(* IEC 61131-3 sources: sceptre-phenix-topologies/cherrymountain-brewery/plant/generated/fleet/fr/openplc/fr-plc-cellar, 1 file *)

(* ---- located_vars.st ---- *)
(* Generated by plantgen from plant/plant.yaml and plant/sites.yaml (site fr). Do not edit. *)
(* Analog values are raw registers: engineering value = raw / 10^scaling. *)
(* RIO I/O is at %IX100.0 / %QX100.0 / %IW100 / %QW100 (v3 and v4 alike). *)
(* PLC memory: bits from %QX0.0 (coils), words from %MW0 (holding register qw_count and up, see modbus_slave.json). *)
VAR
  CEL_CLK_KI01_PV AT %IW100 : UINT; (* Cellar simulation clock (compressed fermentation time), h, x10 *)
  CEL_FV101_TT01_PV AT %IW101 : UINT; (* FV-101 side temperature, degF, x100 *)
  CEL_FV101_TT01_ALM_DEVIATION AT %QX0.0 : BOOL; (* FV-101 side temperature: deviation alarm (high) *)
  CEL_FV101_TT01_ALM_HIGH AT %QX0.1 : BOOL; (* FV-101 side temperature: high alarm (medium) *)
  CEL_FV101_TV01_CMD AT %QX100.0 : BOOL; (* FV-101 side glycol valve command *)
  CEL_FV101_TT02_PV AT %IW102 : UINT; (* FV-101 cone temperature, degF, x100 *)
  CEL_FV101_TT02_ALM_DEVIATION AT %QX0.2 : BOOL; (* FV-101 cone temperature: deviation alarm (medium) *)
  CEL_FV101_TV02_CMD AT %QX100.1 : BOOL; (* FV-101 cone glycol valve command *)
  CEL_FV101_PT01_PV AT %IW103 : UINT; (* FV-101 head pressure (absolute), psia, x100 *)
  CEL_FV101_PT01_ALM_HIGH AT %QX0.3 : BOOL; (* FV-101 head pressure (absolute): high alarm (high) *)
  CEL_FV101_PT01_ALM_LOW AT %QX0.4 : BOOL; (* FV-101 head pressure (absolute): low alarm (low) *)
  CEL_FV101_DT01_PV AT %IW104 : UINT; (* FV-101 apparent extract (sample-port density meter), degP, x100 *)
  CEL_FV101_PCV01_SP AT %QW100 : UINT; (* FV-101 spunding valve setpoint (absolute), psia, x100 *)
  CEL_FV101_ZSO01_PV AT %IX100.0 : BOOL; (* FV-101 spunding valve open (venting) *)
  CEL_FV101_TT01_SP AT %MW0 : UINT; (* FV-101 side temperature setpoint, degF, x100 *)
  CEL_FV101_TT02_SP AT %MW1 : UINT; (* FV-101 cone temperature setpoint, degF, x100 *)
  CEL_FV102_TT01_PV AT %IW105 : UINT; (* FV-102 side temperature, degF, x100 *)
  CEL_FV102_TT01_ALM_DEVIATION AT %QX0.5 : BOOL; (* FV-102 side temperature: deviation alarm (high) *)
  CEL_FV102_TT01_ALM_HIGH AT %QX0.6 : BOOL; (* FV-102 side temperature: high alarm (medium) *)
  CEL_FV102_TV01_CMD AT %QX100.2 : BOOL; (* FV-102 side glycol valve command *)
  CEL_FV102_TT02_PV AT %IW106 : UINT; (* FV-102 cone temperature, degF, x100 *)
  CEL_FV102_TT02_ALM_DEVIATION AT %QX0.7 : BOOL; (* FV-102 cone temperature: deviation alarm (medium) *)
  CEL_FV102_TV02_CMD AT %QX100.3 : BOOL; (* FV-102 cone glycol valve command *)
  CEL_FV102_PT01_PV AT %IW107 : UINT; (* FV-102 head pressure (absolute), psia, x100 *)
  CEL_FV102_PT01_ALM_HIGH AT %QX1.0 : BOOL; (* FV-102 head pressure (absolute): high alarm (high) *)
  CEL_FV102_PT01_ALM_LOW AT %QX1.1 : BOOL; (* FV-102 head pressure (absolute): low alarm (low) *)
  CEL_FV102_DT01_PV AT %IW108 : UINT; (* FV-102 apparent extract (sample-port density meter), degP, x100 *)
  CEL_FV102_PCV01_SP AT %QW101 : UINT; (* FV-102 spunding valve setpoint (absolute), psia, x100 *)
  CEL_FV102_ZSO01_PV AT %IX100.1 : BOOL; (* FV-102 spunding valve open (venting) *)
  CEL_FV102_TT01_SP AT %MW2 : UINT; (* FV-102 side temperature setpoint, degF, x100 *)
  CEL_FV102_TT02_SP AT %MW3 : UINT; (* FV-102 cone temperature setpoint, degF, x100 *)
  CEL_FV103_TT01_PV AT %IW109 : UINT; (* FV-103 side temperature, degF, x100 *)
  CEL_FV103_TT01_ALM_DEVIATION AT %QX1.2 : BOOL; (* FV-103 side temperature: deviation alarm (high) *)
  CEL_FV103_TT01_ALM_HIGH AT %QX1.3 : BOOL; (* FV-103 side temperature: high alarm (medium) *)
  CEL_FV103_TV01_CMD AT %QX100.4 : BOOL; (* FV-103 side glycol valve command *)
  CEL_FV103_TT02_PV AT %IW110 : UINT; (* FV-103 cone temperature, degF, x100 *)
  CEL_FV103_TT02_ALM_DEVIATION AT %QX1.4 : BOOL; (* FV-103 cone temperature: deviation alarm (medium) *)
  CEL_FV103_TV02_CMD AT %QX100.5 : BOOL; (* FV-103 cone glycol valve command *)
  CEL_FV103_PT01_PV AT %IW111 : UINT; (* FV-103 head pressure (absolute), psia, x100 *)
  CEL_FV103_PT01_ALM_HIGH AT %QX1.5 : BOOL; (* FV-103 head pressure (absolute): high alarm (high) *)
  CEL_FV103_PT01_ALM_LOW AT %QX1.6 : BOOL; (* FV-103 head pressure (absolute): low alarm (low) *)
  CEL_FV103_DT01_PV AT %IW112 : UINT; (* FV-103 apparent extract (sample-port density meter), degP, x100 *)
  CEL_FV103_PCV01_SP AT %QW102 : UINT; (* FV-103 spunding valve setpoint (absolute), psia, x100 *)
  CEL_FV103_ZSO01_PV AT %IX100.2 : BOOL; (* FV-103 spunding valve open (venting) *)
  CEL_FV103_TT01_SP AT %MW4 : UINT; (* FV-103 side temperature setpoint, degF, x100 *)
  CEL_FV103_TT02_SP AT %MW5 : UINT; (* FV-103 cone temperature setpoint, degF, x100 *)
  CEL_FV104_TT01_PV AT %IW113 : UINT; (* FV-104 side temperature, degF, x100 *)
  CEL_FV104_TT01_ALM_DEVIATION AT %QX1.7 : BOOL; (* FV-104 side temperature: deviation alarm (high) *)
  CEL_FV104_TT01_ALM_HIGH AT %QX2.0 : BOOL; (* FV-104 side temperature: high alarm (medium) *)
  CEL_FV104_TV01_CMD AT %QX100.6 : BOOL; (* FV-104 side glycol valve command *)
  CEL_FV104_TT02_PV AT %IW114 : UINT; (* FV-104 cone temperature, degF, x100 *)
  CEL_FV104_TT02_ALM_DEVIATION AT %QX2.1 : BOOL; (* FV-104 cone temperature: deviation alarm (medium) *)
  CEL_FV104_TV02_CMD AT %QX100.7 : BOOL; (* FV-104 cone glycol valve command *)
  CEL_FV104_PT01_PV AT %IW115 : UINT; (* FV-104 head pressure (absolute), psia, x100 *)
  CEL_FV104_PT01_ALM_HIGH AT %QX2.2 : BOOL; (* FV-104 head pressure (absolute): high alarm (high) *)
  CEL_FV104_PT01_ALM_LOW AT %QX2.3 : BOOL; (* FV-104 head pressure (absolute): low alarm (low) *)
  CEL_FV104_DT01_PV AT %IW116 : UINT; (* FV-104 apparent extract (sample-port density meter), degP, x100 *)
  CEL_FV104_PCV01_SP AT %QW103 : UINT; (* FV-104 spunding valve setpoint (absolute), psia, x100 *)
  CEL_FV104_ZSO01_PV AT %IX100.3 : BOOL; (* FV-104 spunding valve open (venting) *)
  CEL_FV104_TT01_SP AT %MW6 : UINT; (* FV-104 side temperature setpoint, degF, x100 *)
  CEL_FV104_TT02_SP AT %MW7 : UINT; (* FV-104 cone temperature setpoint, degF, x100 *)
  CEL_BBT201_TT01_PV AT %IW117 : UINT; (* BBT-201 temperature, degF, x100 *)
  CEL_BBT201_TT01_ALM_DEVIATION AT %QX2.4 : BOOL; (* BBT-201 temperature: deviation alarm (medium) *)
  CEL_BBT201_PT01_PV AT %IW118 : UINT; (* BBT-201 head pressure (absolute), psia, x100 *)
  CEL_BBT201_PT01_ALM_HIGH AT %QX2.5 : BOOL; (* BBT-201 head pressure (absolute): high alarm (high) *)
  CEL_BBT201_LT01_PV AT %IW119 : UINT; (* BBT-201 level, %, x10 *)
  CEL_BBT201_AT01_PV AT %IW120 : UINT; (* BBT-201 dissolved CO2 (inline meter), vol, x100 *)
  CEL_BBT201_FT01_PV AT %IW121 : UINT; (* BBT-201 carbonation stone CO2 flow, L/min, x10 *)
  CEL_BBT201_TV01_CMD AT %QX101.0 : BOOL; (* BBT-201 jacket glycol valve command *)
  CEL_BBT201_XV01_CMD AT %QX101.1 : BOOL; (* BBT-201 outlet valve (to packaging) *)
  CEL_BBT201_FCV01_OUT AT %QW104 : UINT; (* BBT-201 carbonation CO2 flow valve position, %, x10 *)
  CEL_BBT201_TT01_SP AT %MW8 : UINT; (* BBT-201 temperature setpoint, degF, x100 *)
  CEL_BBT201_AT01_SP AT %MW9 : UINT; (* BBT-201 carbonation target, vol, x100 *)
  CEL_BBT201_PT01_SP AT %MW10 : UINT; (* BBT-201 equilibrium head pressure for the target (computed, absolute), psia, x100 *)
  CEL_BBT202_TT01_PV AT %IW122 : UINT; (* BBT-202 temperature, degF, x100 *)
  CEL_BBT202_TT01_ALM_DEVIATION AT %QX2.6 : BOOL; (* BBT-202 temperature: deviation alarm (medium) *)
  CEL_BBT202_PT01_PV AT %IW123 : UINT; (* BBT-202 head pressure (absolute), psia, x100 *)
  CEL_BBT202_PT01_ALM_HIGH AT %QX2.7 : BOOL; (* BBT-202 head pressure (absolute): high alarm (high) *)
  CEL_BBT202_LT01_PV AT %IW124 : UINT; (* BBT-202 level, %, x10 *)
  CEL_BBT202_AT01_PV AT %IW125 : UINT; (* BBT-202 dissolved CO2 (inline meter), vol, x100 *)
  CEL_BBT202_FT01_PV AT %IW126 : UINT; (* BBT-202 carbonation stone CO2 flow, L/min, x10 *)
  CEL_BBT202_TV01_CMD AT %QX101.2 : BOOL; (* BBT-202 jacket glycol valve command *)
  CEL_BBT202_XV01_CMD AT %QX101.3 : BOOL; (* BBT-202 outlet valve (to packaging) *)
  CEL_BBT202_FCV01_OUT AT %QW105 : UINT; (* BBT-202 carbonation CO2 flow valve position, %, x10 *)
  CEL_BBT202_TT01_SP AT %MW11 : UINT; (* BBT-202 temperature setpoint, degF, x100 *)
  CEL_BBT202_AT01_SP AT %MW12 : UINT; (* BBT-202 carbonation target, vol, x100 *)
  CEL_BBT202_PT01_SP AT %MW13 : UINT; (* BBT-202 equilibrium head pressure for the target (computed, absolute), psia, x100 *)
  CEL_DH_ZSC01_PV AT %IX100.4 : BOOL; (* Hop port closed *)
  CEL_DH_XV01_CMD AT %QX101.4 : BOOL; (* Hop port CO2 purge valve *)
  CEL_DH_XV02_CMD AT %QX101.5 : BOOL; (* Hop dose valve *)
  CEL_DH_XC01_CMD AT %QX3.0 : BOOL; (* Dry-hop dose request (operator; fr-plc-cellar purges, doses, and clears it) *)
  CEL_DH_XS01_STEP AT %MW14 : UINT; (* Dry-hop sequence step (0 idle, 1 CO2 purge, 2 dose), None, x1 *)
  CEL_XFER_ZS01_PV AT %IX100.5 : BOOL; (* Transfer route verified (swing-panel proximity) *)
  CEL_XFER_YS01_PV AT %IX100.6 : BOOL; (* Transfer pump running *)
  CEL_XFER_FT01_PV AT %IW127 : UINT; (* Transfer flow, gal/min, x10 *)
  CEL_XFER_HS01_CMD AT %QX101.6 : BOOL; (* Transfer pump run command *)
  CEL_XFER_XS01_ACTIVE AT %QX3.1 : BOOL; (* Transfer in progress (peer status for fr-plc-utilities) *)
  CEL_XFER_XS02_CIP_PERMIT AT %QX3.2 : BOOL; (* CIP permitted on the cellar circuits (peer status for fr-plc-utilities) *)
  CEL_SYS_XS01_CO2_OK AT %IX100.7 : BOOL; (* Cellar CO2 relay healthy (below 15,000 ppm, detection powered) *)
  CEL_SYS_XS01_CO2_INHIBIT AT %QX3.3 : BOOL; (* Carbonation inhibited by the cellar CO2 relay (fr-plc-cellar interlock) *)
  CEL_SYS_XS01_ALM_STATE AT %QX3.4 : BOOL; (* Carbonation inhibited by the cellar CO2 relay (fr-plc-cellar interlock): state alarm (medium) *)
  CEL_PSV_ZSH01_PV AT %IX101.0 : BOOL; (* FV-101 relief valve (PSV) lifted *)
  CEL_PSV_ZSH01_ALM_STATE AT %QX3.5 : BOOL; (* FV-101 relief valve (PSV) lifted: state alarm (high) *)
  CEL_PSV_ZSH02_PV AT %IX101.1 : BOOL; (* FV-102 relief valve (PSV) lifted *)
  CEL_PSV_ZSH02_ALM_STATE AT %QX3.6 : BOOL; (* FV-102 relief valve (PSV) lifted: state alarm (high) *)
  CEL_PSV_ZSH03_PV AT %IX101.2 : BOOL; (* FV-103 relief valve (PSV) lifted *)
  CEL_PSV_ZSH03_ALM_STATE AT %QX3.7 : BOOL; (* FV-103 relief valve (PSV) lifted: state alarm (high) *)
  CEL_PSV_ZSH04_PV AT %IX101.3 : BOOL; (* FV-104 relief valve (PSV) lifted *)
  CEL_PSV_ZSH04_ALM_STATE AT %QX4.0 : BOOL; (* FV-104 relief valve (PSV) lifted: state alarm (high) *)
  CEL_PSV_ZSH05_PV AT %IX101.4 : BOOL; (* BBT-201 relief valve (PSV) lifted *)
  CEL_PSV_ZSH05_ALM_STATE AT %QX4.1 : BOOL; (* BBT-201 relief valve (PSV) lifted: state alarm (high) *)
  CEL_PSV_ZSH06_PV AT %IX101.5 : BOOL; (* BBT-202 relief valve (PSV) lifted *)
  CEL_PSV_ZSH06_ALM_STATE AT %QX4.2 : BOOL; (* BBT-202 relief valve (PSV) lifted: state alarm (high) *)
  CEL_ENTRY_HS01_ENTRY AT %QX4.3 : BOOL; (* FV-101 entry permit issued (entry supervisor; locks the vessel out) *)
  CEL_ENTRY_HS02_ENTRY AT %QX4.4 : BOOL; (* FV-102 entry permit issued (entry supervisor; locks the vessel out) *)
  CEL_ENTRY_HS03_ENTRY AT %QX4.5 : BOOL; (* FV-103 entry permit issued (entry supervisor; locks the vessel out) *)
  CEL_ENTRY_HS04_ENTRY AT %QX4.6 : BOOL; (* FV-104 entry permit issued (entry supervisor; locks the vessel out) *)
  CEL_ENTRY_HS05_ENTRY AT %QX4.7 : BOOL; (* BBT-201 entry permit issued (entry supervisor; locks the vessel out) *)
  CEL_ENTRY_HS06_ENTRY AT %QX5.0 : BOOL; (* BBT-202 entry permit issued (entry supervisor; locks the vessel out) *)
  CEL_ENTRY_XS01_LOCKED AT %QX5.1 : BOOL; (* FV-101 locked out for entry (glycol, CO2, outlet, and CIP) *)
  CEL_ENTRY_XS02_LOCKED AT %QX5.2 : BOOL; (* FV-102 locked out for entry (glycol, CO2, outlet, and CIP) *)
  CEL_ENTRY_XS03_LOCKED AT %QX5.3 : BOOL; (* FV-103 locked out for entry (glycol, CO2, outlet, and CIP) *)
  CEL_ENTRY_XS04_LOCKED AT %QX5.4 : BOOL; (* FV-104 locked out for entry (glycol, CO2, outlet, and CIP) *)
  CEL_ENTRY_XS05_LOCKED AT %QX5.5 : BOOL; (* BBT-201 locked out for entry (glycol, CO2, outlet, and CIP) *)
  CEL_ENTRY_XS06_LOCKED AT %QX5.6 : BOOL; (* BBT-202 locked out for entry (glycol, CO2, outlet, and CIP) *)
  CEL_ENTRY_XS11_CIP_OK AT %QX5.7 : BOOL; (* FV-101 CIP permitted, not in entry (peer status for fr-plc-utilities) *)
  CEL_ENTRY_XS12_CIP_OK AT %QX6.0 : BOOL; (* FV-102 CIP permitted, not in entry (peer status for fr-plc-utilities) *)
  CEL_ENTRY_XS13_CIP_OK AT %QX6.1 : BOOL; (* FV-103 CIP permitted, not in entry (peer status for fr-plc-utilities) *)
  CEL_ENTRY_XS14_CIP_OK AT %QX6.2 : BOOL; (* FV-104 CIP permitted, not in entry (peer status for fr-plc-utilities) *)
  CEL_ENTRY_XS15_CIP_OK AT %QX6.3 : BOOL; (* BBT-201 CIP permitted, not in entry (peer status for fr-plc-utilities) *)
  CEL_ENTRY_XS16_CIP_OK AT %QX6.4 : BOOL; (* BBT-202 CIP permitted, not in entry (peer status for fr-plc-utilities) *)
  CEL_ENTRY_XA01_PV AT %QX6.5 : BOOL; (* FV-101 write to a locked-out valve during entry *)
  CEL_ENTRY_XA01_ALM_STATE AT %QX6.6 : BOOL; (* FV-101 write to a locked-out valve during entry: state alarm (critical) *)
  CEL_ENTRY_XA02_PV AT %QX6.7 : BOOL; (* FV-102 write to a locked-out valve during entry *)
  CEL_ENTRY_XA02_ALM_STATE AT %QX7.0 : BOOL; (* FV-102 write to a locked-out valve during entry: state alarm (critical) *)
  CEL_ENTRY_XA03_PV AT %QX7.1 : BOOL; (* FV-103 write to a locked-out valve during entry *)
  CEL_ENTRY_XA03_ALM_STATE AT %QX7.2 : BOOL; (* FV-103 write to a locked-out valve during entry: state alarm (critical) *)
  CEL_ENTRY_XA04_PV AT %QX7.3 : BOOL; (* FV-104 write to a locked-out valve during entry *)
  CEL_ENTRY_XA04_ALM_STATE AT %QX7.4 : BOOL; (* FV-104 write to a locked-out valve during entry: state alarm (critical) *)
  CEL_ENTRY_XA05_PV AT %QX7.5 : BOOL; (* BBT-201 write to a locked-out valve during entry *)
  CEL_ENTRY_XA05_ALM_STATE AT %QX7.6 : BOOL; (* BBT-201 write to a locked-out valve during entry: state alarm (critical) *)
  CEL_ENTRY_XA06_PV AT %QX7.7 : BOOL; (* BBT-202 write to a locked-out valve during entry *)
  CEL_ENTRY_XA06_ALM_STATE AT %QX8.0 : BOOL; (* BBT-202 write to a locked-out valve during entry: state alarm (critical) *)
  CEL_PROFILE_HS01_AUTO AT %QX8.1 : BOOL; (* FV-101 fermentation profile on (fr-plc-cellar sets its temperature setpoints) *)
  CEL_PROFILE_HS02_AUTO AT %QX8.2 : BOOL; (* FV-102 fermentation profile on (fr-plc-cellar sets its temperature setpoints) *)
  CEL_PROFILE_HS03_AUTO AT %QX8.3 : BOOL; (* FV-103 fermentation profile on (fr-plc-cellar sets its temperature setpoints) *)
  CEL_PROFILE_HS04_AUTO AT %QX8.4 : BOOL; (* FV-104 fermentation profile on (fr-plc-cellar sets its temperature setpoints) *)
  CEL_PROFILE_KS01_STAGE AT %MW15 : UINT; (* FV-101 profile stage (0 empty, 1 fermenting, 2 diacetyl rest, 3 crash), None, x1 *)
  CEL_PROFILE_KS02_STAGE AT %MW16 : UINT; (* FV-102 profile stage (0 empty, 1 fermenting, 2 diacetyl rest, 3 crash), None, x1 *)
  CEL_PROFILE_KS03_STAGE AT %MW17 : UINT; (* FV-103 profile stage (0 empty, 1 fermenting, 2 diacetyl rest, 3 crash), None, x1 *)
  CEL_PROFILE_KS04_STAGE AT %MW18 : UINT; (* FV-104 profile stage (0 empty, 1 fermenting, 2 diacetyl rest, 3 crash), None, x1 *)
  CEL_PROFILE_TC01_SP AT %MW19 : UINT; (* Profile temperature while the beer ferments, degF, x100 *)
  CEL_PROFILE_TC02_SP AT %MW20 : UINT; (* Profile temperature of the diacetyl rest, degF, x100 *)
  CEL_PROFILE_TC03_SP AT %MW21 : UINT; (* Profile temperature of the crash, degF, x100 *)
  CEL_PROFILE_KC01_SP AT %MW22 : UINT; (* Diacetyl rest length in plant minutes (180 is 144 h of fermentation on the range's 48x clock), min, x1 *)
END_VAR
